ABB RAPID module: DropOut1.mod

%%%
  VERSION:1
  LANGUAGE:ENGLISH
%%%
MODULE MOD_DropOut1

    ! -------------------------------
    ! Define customized variables here
    ! ...

	! Tool variables:
	PERS tooldata SuctionCup := [TRUE,[[-94.709,0.000,259.352],[0.00000000,0.00000000,0.00000000,1.00000000]],[1,[0,0,20],[1,0,0,0],0,0,0.005]];

	! Reference variables:
	PERS wobjdata Out := [FALSE, TRUE, "", [[0,0,0],[1,0,0,0]],[[290.000,-450.000,10.000],[1.00000000,0.00000000,0.00000000,0.00000000]]];

	PROC Main()
		ConfJ \On;
		ConfL \Off;
		! Program generated by VerticalBot Studio for ABB IRB 1200-5/0.9 on 25/10/2026 12:00:00
		! Using nominal kinematics.
		MoveAbsJ [[-66.056500,21.575200,36.080800,0.000000,32.344000,-66.056500],[9E+09,9E+09,9E+09,9E+09,9E+09,9E+09]],v500,z1,SuctionCup \WObj:=Out;
		MoveL [[-16.111,46.392,30.000],[0.00000000,1.00000000,0.00000000,-0.00000000],[-1,0,-1,0],[9E+09,9E+09,9E+09,9E+09,9E+09,9E+09]],v500,z1,SuctionCup \WObj:=Out;
		! Detach from Suction Cup
		WaitTime 0.500;
		MoveL [[-16.111,46.485,105.701],[0.00000000,1.00000000,0.00000000,-0.00000000],[-1,0,-1,0],[9E+09,9E+09,9E+09,9E+09,9E+09,9E+09]],v500,z1,SuctionCup \WObj:=Out;
	ENDPROC

ENDMODULE
